(* PLC project sfc_batch_fill_drain_bomb, Anonymous Benchmark Suite 1.0 *)
(* stored: creationDateTime 2026-08-26T00:00:00 *)

PROGRAM batch_cycle
  VAR_INPUT
    start : BOOL;
    level_high : BOOL;
    reaction_done : BOOL;
    level_low : BOOL;
  END_VAR
  VAR_OUTPUT
    fill_valve : BOOL;
    drain_valve : BOOL;
  END_VAR

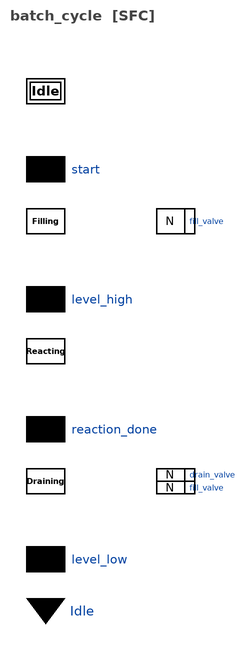
INITIAL_STEP Idle:
END_STEP
TRANSITION FROM Idle TO Filling
  := start;
END_TRANSITION
STEP Filling:
  fill_valve(N);
END_STEP
TRANSITION FROM Filling TO Reacting
  := level_high;
END_TRANSITION
STEP Reacting:
END_STEP
TRANSITION FROM Reacting TO Draining
  := reaction_done;
END_TRANSITION
STEP Draining:
  drain_valve(N);
  fill_valve(N);
END_STEP
TRANSITION FROM Draining TO Idle
  := level_low;
END_TRANSITION
END_PROGRAM

CONFIGURATION Config0
  RESOURCE Res0 ON PLC
    TASK tcyclic(INTERVAL := T#10ms, PRIORITY := 0);
    PROGRAM inst0 WITH tcyclic : batch_cycle;
  END_RESOURCE
END_CONFIGURATION
